// Mitsubishi GX Works2 project: Task_3_Ex2   PLC: FX3G

PROGRAM MAIN
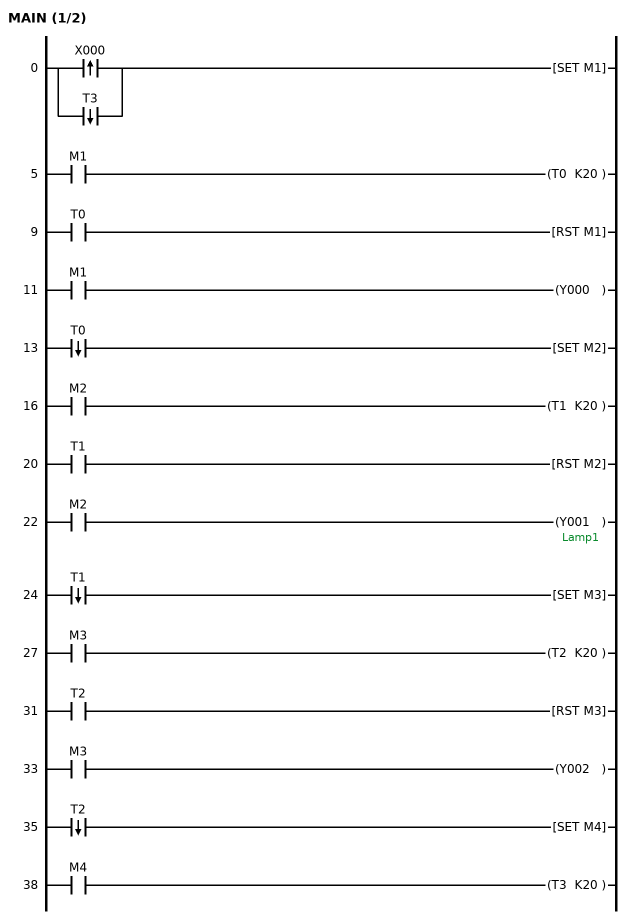
0     LDP     X000
      ORF     T3
      SET     M1
5     LD      M1
      OUT     T0 K20
9     LD      T0
      RST     M1
11    LD      M1
      OUT     Y000
13    LDF     T0
      SET     M2
16    LD      M2
      OUT     T1 K20
20    LD      T1
      RST     M2
22    LD      M2
      OUT     Y001  ; Lamp1
24    LDF     T1
      SET     M3
27    LD      M3
      OUT     T2 K20
31    LD      T2
      RST     M3
33    LD      M3
      OUT     Y002
35    LDF     T2
      SET     M4
38    LD      M4
      OUT     T3 K20
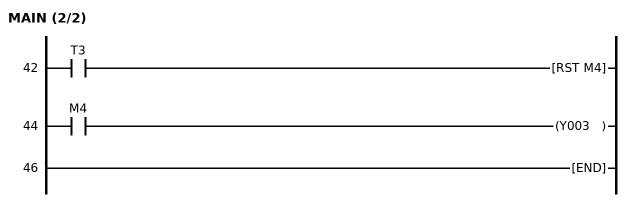
42    LD      T3
      RST     M4
44    LD      M4
      OUT     Y003
46    END
END_PROGRAM
